Fanuc KAREL source: ks00054.KL

-- PROVISIONAL review KL for V770-1; original PC SHA256 41dc8e2b7a7dd04336e4914824e0288dfbc50e9edf2ace4daf9276526e2bd691
-- Incomplete behavior may be omitted. Consult companion uncertainty JSON. Do not deploy.
PROGRAM KS00054
%NOLOCKGROUP
BEGIN
  -- UNRESOLVED_PC offsets 5-13; opcodes 3F,75
  -- UNRESOLVED_PC offsets 18-27; opcodes 3F,75
  -- UNRESOLVED_PC offsets 32-45; opcodes 22,1D,23
  -- UNRESOLVED_PC offsets 50-54; opcodes 7F
END KS00054
